StartTest(TestName := 'Test_TriggerForOneCycleOnRisingEdge');
group_1(Run := TRUE, ErrAck := FALSE); // T_SafeGroup
fb_1(Signal := FALSE); // T_SafeRTrig_UserFB
AssertEquals_BOOL(Expected := FALSE, Actual := fb_1.Trigger, Message := 'no trigger while the signal is off');
fb_1(Signal := TRUE); // T_SafeRTrig_UserFB
AssertEquals_BOOL(Expected := TRUE, Actual := fb_1.Trigger, Message := 'trigger on the rising edge');
fb_1(Signal := TRUE); // T_SafeRTrig_UserFB
AssertEquals_BOOL(Expected := FALSE, Actual := fb_1.Trigger, Message := 'trigger lasts one cycle');
fb_1(Signal := FALSE); // T_SafeRTrig_UserFB
AssertEquals_BOOL(Expected := FALSE, Actual := fb_1.Trigger, Message := 'no trigger on the falling edge');
fb_1(Signal := TRUE); // T_SafeRTrig_UserFB
AssertEquals_BOOL(Expected := TRUE, Actual := fb_1.Trigger, Message := 'triggers again on the next rising edge');
FinishTest(TestName := 'Test_TriggerForOneCycleOnRisingEdge');
END_METHOD

END_FUNCTION_BLOCK

// ---- Examples/PRG_EStopExample.TcPOU
// Worked example: a two-channel emergency stop with contactor feedback, wired the way a
// TwinSAFE project links it, plus the standard PLC signals (Run, ErrAck, Restart).
// The blocks join the group at declaration; call the group before its members.
// Toggle the "field" variables online to trial the behaviour and watch the State / Diag outputs.
PROGRAM PRG_EStopExample
VAR
    // --- simulated field devices (real hardware in a TwinSAFE system)
    eStopChannel1 : BOOL := TRUE; // NC contact, TRUE = not pressed
    eStopChannel2 : BOOL := TRUE;

    // --- standard PLC interface to the TwinSAFE group (linked to standard variables)
    safetyRun : BOOL := TRUE;
    safetyErrAck : BOOL;
    restartButton : BOOL; // 0 -> 1 -> 0 to restart

    // --- TwinSAFE model: the group, then its members (parameters as in the Safety Editor property grid)
    group : T_SafeGroup;
    inputTerminal : T_SafeInputTerminal(group := group); // EL1904
    outputTerminal : T_SafeOutputTerminal(group := group); // EL2904
    eStop : T_SafeEStop(group := group) := (Parameters := (DiscrepancyTime1 := T#500MS, DelayTime := T#1S));

    // --- simulated contactors: pull in 50 ms after the safe output energises; EDM1 = NOT pulled in
    contactorPullIn : TON;
END_VAR

// TwinSAFE group: standard PLC signals in; it reads its members' states itself
group(Run := safetyRun, ErrAck := safetyErrAck);

// Field -> safe input terminal (EL1904)
inputTerminal(Channel1 := eStopChannel1, Channel2 := eStopChannel2);

// FB ESTOP wired as in the safety project: EStopIn1/2 two channel, EDM1 and Restart from standard signals
eStop(
    Restart := restartButton,
    EDM1 := NOT contactorPullIn.Q,
    EStopIn1 := inputTerminal.SafeIn1,
    EStopIn2 := inputTerminal.SafeIn2
);

// Safe outputs -> output terminal (EL2904) -> field
outputTerminal(SafeOut1 := eStop.EStopOut, SafeOut2 := eStop.EStopDelOut);

// Simulated contactors follow the field output
contactorPullIn(IN := outputTerminal.Channel1, PT := T#50MS);

END_PROGRAM

// ---- Core/T_SafeOutputTerminal.TcPOU
// Model of a four channel safe output terminal (EL2904): a TwinSAFE connection with four channels.
// Declare it in its group:  outputTerminal : T_SafeOutputTerminal(group := safetyGroup);
// SafeOut1..4 are wired from FB outputs; Channel1..4 are the simulated field outputs,
// forced FALSE (fail-safe) unless the connection is in the Data state and the group is in RUN (OutputsEnabled).
FUNCTION_BLOCK T_SafeOutputTerminal EXTENDS T_SafeConnection
VAR_INPUT
    SafeOut1 : BOOL;
    SafeOut2 : BOOL;
    SafeOut3 : BOOL;
    SafeOut4 : BOOL;
END_VAR
VAR_OUTPUT
    Channel1 : BOOL;
    Channel2 : BOOL;
    Channel3 : BOOL;
    Channel4 : BOOL;
END_VAR

SUPER^();
Channel1 := SafeOut1 AND OutputsEnabled;
Channel2 := SafeOut2 AND OutputsEnabled;
Channel3 := SafeOut3 AND OutputsEnabled;
Channel4 := SafeOut4 AND OutputsEnabled;

END_FUNCTION_BLOCK

// ---- Examples/PRG_EStopExample_CFC.TcPOU
// Worked example: a two-channel emergency stop with contactor feedback, wired the way a
// TwinSAFE project links it, plus the standard PLC signals (Run, ErrAck, Restart).
// The blocks join the group at declaration; call the group before its members.
// CFC twin of PRG_EStopExample: the same wiring as a diagram.
// Toggle the "field" variables online to trial the behaviour and watch the State / Diag outputs.
PROGRAM PRG_EStopExample_CFC
VAR
    // --- simulated field devices (real hardware in a TwinSAFE system)
    eStopChannel1 : BOOL := TRUE; // NC contact, TRUE = not pressed
    eStopChannel2 : BOOL := TRUE;

    // --- standard PLC interface to the TwinSAFE group (linked to standard variables)
    safetyRun : BOOL := TRUE;
    safetyErrAck : BOOL;
    restartButton : BOOL; // 0 -> 1 -> 0 to restart

    // --- TwinSAFE model: the group, then its members (parameters as in the Safety Editor property grid)
    group : T_SafeGroup;
    inputTerminal : T_SafeInputTerminal(group := group); // EL1904
    outputTerminal : T_SafeOutputTerminal(group := group); // EL2904
    eStop : T_SafeEStop(group := group) := (Parameters := (DiscrepancyTime1 := T#500MS, DelayTime := T#1S));

    // --- simulated contactors: pull in 50 ms after the safe output energises; EDM1 = NOT pulled in
    contactorPullIn : TON;
END_VAR

group(Run := safetyRun, ErrAck := safetyErrAck); // T_SafeGroup
contactorPullIn(IN := outputTerminal.Channel1, PT := T#50MS); // TON
inputTerminal(Channel1 := eStopChannel1, Channel2 := eStopChannel2); // T_SafeInputTerminal
eStop(
    Restart := restartButton,
    EDM1 := NOT contactorPullIn.Q,
    EStopIn1 := inputTerminal.SafeIn1,
    EStopIn2 := inputTerminal.SafeIn2); // T_SafeEStop
outputTerminal(SafeOut1 := eStop.EStopOut, SafeOut2 := eStop.EStopDelOut); // T_SafeOutputTerminal

END_PROGRAM

// ---- Project Information/F_GetCompany.TcPOU
// This function has been automatically generated from the project information.
{attribute 'signature_flag' := '1073741824'}
{attribute 'TcGenerated'}
{attribute 'no-analysis'}
FUNCTION F_GetCompany : WSTRING
VAR_INPUT
	
END_VAR

F_GetCompany := "Intecre Ltd";

END_FUNCTION

// ---- Project Information/F_GetTitle.TcPOU
// This function has been automatically generated from the project information.
{attribute 'signature_flag' := '1073741824'}
{attribute 'TcGenerated'}
{attribute 'no-analysis'}
FUNCTION F_GetTitle : WSTRING
VAR_INPUT
	
END_VAR

F_GetTitle := "Intecre.TwinSAFE.Models";

END_FUNCTION

// ---- Project Information/F_GetVersion.TcPOU
// This function has been automatically generated from the project information.
{attribute 'signature_flag' := '1073741824'}
{attribute 'TcGenerated'}
{attribute 'no-analysis'}
FUNCTION F_GetVersion : ST_LibVersion
VAR_INPUT
	
END_VAR

F_GetVersion.iMajor := 0;
F_GetVersion.iMinor := 5;
F_GetVersion.iBuild := 0;
F_GetVersion.iRevision := 3;
F_GetVersion.sVersion := '0.5.0.3';
F_GetVersion.nFlags := 0;

END_FUNCTION
